FUNCTION_BLOCK FB_DomeClosingState EXTENDS  FB_DomeState
VAR
	Stage		: UINT:= 0;
	tonSleep	: TON := (PT:=T#5S);
	tonTimeout	: TON:= (PT:=T#3M); // see Baader Handbook
	// #202: d#closhut is acknowledged (d#gotmess) but the shutter stays open (d#shutope): the command is sent again at
	// most nMaxAttempts times in all, then it is an error. Before, it was sent for ever, because the timeout is stopped
	// at every poll, and nothing was logged.
	nAttempts	: UINT;
	nMaxAttempts: UINT := 3;
END_VAR


METHOD CloseCommand : BOOL
// #202: a new close starts the shutter command again, with a fresh count
LogEvent(sText := 'Dome: close received while closing, the shutter command is started again', sLevel := 'WARNING');
nAttempts := 0;
Stage := 0;
tonSleep(IN:=FALSE);
tonTimeout(IN:=FALSE);
END_METHOD

METHOD FoundError : BOOL
nAttempts := 0;
Stage:= 0;
tonSleep(IN:=FALSE);
tonTimeout(IN:=FALSE);
pDome^._Error := TRUE;
pDome^.SetState(pDome^.fbDomeErrorState);
END_METHOD


METHOD OpenCommand : BOOL
nAttempts := 0;
Stage:= 0;
tonSleep(IN:=FALSE);
tonTimeout(IN:=FALSE);
pDome^.SetState(pDome^.fbDomeOpeningState);
END_METHOD

METHOD RunState : BOOL
VAR_INPUT
END_VAR
CASE Stage OF
	0:
		tonTimeout(IN:=TRUE);
		Stage := 1;
	1:
		pDome^.fbSend(	SendString:= 'd#closhut',
					TXbuffer:= TxBufferDome,
					Busy=>,
					Error=> );
		IF NOT pDome^.fbSend.Busy  THEN
			Stage := 2;
		END_IF
	2:
		IF pDome^.bStringReceived THEN
			IF pDome^._ReceivedString = 'd#comerro' OR pDome^._ReceivedString = 'd#domerro' THEN
				foundError();
			ELSIF pDome^._ReceivedString = 'd#gotmess' THEN
				Stage := 3;
			END_IF
		ELSIF NOT pDome^.fbReceive.Busy THEN
			tonSleep(IN:=TRUE);
			IF tonSleep.Q THEN
				tonSleep(IN:=FALSE);
				Stage := 1;
			END_IF
		END_IF
		tonTimeout(IN:=TRUE);
		IF tonTimeout.Q THEN
			tonTimeout(IN:=FALSE);
			foundError();
		END_IF
	3:
		tonTimeout(IN:=FALSE);
		
		tonSleep(IN:=TRUE);
		IF tonSleep.Q THEN
			tonSleep(IN:=FALSE);
			Stage := 4;
			tonTimeout(IN:=TRUE);
		END_IF
	4:
		pDome^.fbSend(	SendString:= 'd#getshut',
					TXbuffer:= TxBufferDome,
					Busy=>,
					Error=> );
		IF NOT pDome^.fbSend.Busy  THEN
			Stage := 5;
		END_IF
	5: 
		IF pDome^.bStringReceived THEN
			IF pDome^._ReceivedString = 'd#comerro' OR pDome^._ReceivedString = 'd#domerro' THEN
				FoundError();
			ELSIF pDome^._ReceivedString = 'd#shutclo' THEN
				pDome^._DomeShutterState := E_RoofState.closed;
				Stage := 6;
			ELSIF pDome^._ReceivedString = 'd#shutope' THEN
				pDome^._DomeShutterState := E_RoofState.opened;
				nAttempts := nAttempts + 1;
				IF nAttempts >= nMaxAttempts THEN
					LogEvent(sText := 'Dome: the shutter does not close, d#closhut is acknowledged but the shutter stays open', sLevel := 'WARNING');
					FoundError();
				ELSE
					Stage := 0;
				END_IF
			ELSIF pDome^._ReceivedString = 'd#shutrun' THEN
				pDome^._DomeShutterState := E_RoofState.closing;
				Stage := 3;
			END_IF
		ELSIF NOT pDome^.fbReceive.Busy THEN
			// mixed up string? ask again
			tonSleep(IN:=TRUE);
			IF tonSleep.Q THEN
				tonSleep(IN:=FALSE);
				Stage := 4;
			END_IF
		END_IF
		tonTimeout(IN:=TRUE);
		IF tonTimeout.Q THEN
			tonTimeout(IN:=FALSE);
			FoundError();
		END_IF
	
	6:
		tonTimeout(IN:=FALSE);
		SuccessfulFinished();
		
END_CASE
END_METHOD


PROPERTY StateID : STRING
GET
StateID := 'Closing State';
END_GET
END_PROPERTY


METHOD SuccessfulFinished : BOOL
nAttempts := 0;
Stage:= 0;
tonSleep(IN:=FALSE);
tonTimeout(IN:=FALSE);
pDome^.SetState(pDome^.fbDomeIdleState);
END_METHOD

END_FUNCTION_BLOCK

(* stored: Version 1.1.0.1, ProductVersion 3.1.4024.15
   POU FB_DomeClosingState: Id {8a6f5a3c-ae72-4eae-976a-7d93edd4c94d}, SpecialFunc None
   Method CloseCommand: Id {f429e250-eab4-46cf-960e-227731c324e9}
   Method FoundError: Id {96dff545-3011-469a-a894-b669fe57425f}
   Method OpenCommand: Id {0e03056c-1c74-4cff-8ebd-a639f27039c7}
   Method RunState: Id {90c99c1b-0afb-40a6-bb12-4cc551df7cd1}
   Property StateID: Id {b6536c1f-6c30-4c70-bf10-aba7df39f93f}
   Get Get: Id {190c2a86-afe4-41f2-97fa-37fbda85f6bd}
   Method SuccessfulFinished: Id {065936d6-e0cd-40ab-a52b-24456541a2fb} *)
